Fanuc KAREL source: ka00215.KL

PROGRAM KA00215
%STACKSIZE=65535
%PRIORITY=65535
%NOLOCKGROUP
VAR
SRC : ARRAY[4] OF XYZWPR
DST : ARRAY[4] OF XYZWPR
BEGIN
-- UNRESOLVED_PC line 7 opcodes [22 22 1E] marker_code=0
END KA00215
